(* IEC 61131-3 sources: sis-interlock-demo/src/POUs/Sis/F_VoteArchChannels, 2 files *)

(* ---- F_VoteArchChannels.decl.st ---- *)
// Назначение: число каналов N схемы голосования по таблице 5.1; 0 — для None, ForcedTrip и
//             значений вне перечисления.
// Автор:      kr0nsch
// Версия:     0.1.0
// Документ:   docs/DESIGN.md, раздел «5.10 Вспомогательные функции голосования»
// ВНИМАНИЕ:   код демонстрационный и не предназначен для систем безопасности. Реальная ПАЗ
//             требует определения SIL, сертифицированных аппаратных и программных средств
//             и валидации по ГОСТ Р МЭК 61511.
FUNCTION F_VoteArchChannels : UINT
VAR_INPUT
    eArch : E_VoteArch;   // схема голосования
END_VAR

(* ---- F_VoteArchChannels.impl.st ---- *)
CASE eArch OF
    E_VoteArch.Vote1oo1:
        F_VoteArchChannels := 1;
    E_VoteArch.Vote1oo2, E_VoteArch.Vote2oo2:
        F_VoteArchChannels := 2;
    E_VoteArch.Vote2oo3:
        F_VoteArchChannels := GVL_Const.VOTE_2OO3_CHANNELS;
ELSE
    // None, ForcedTrip и значения вне перечисления — схемы нет
    F_VoteArchChannels := 0;
END_CASE
